// TIA Portal V21 export
// export: Created 2026-11-21T13:31:41.9826464Z, ExportSetting WithDefaults, DisplayName Totally Integrated Automation Portal, DisplayVersion V21, DisplayName STEP 7 Professional, DisplayVersion V21, DisplayName STEP 7 Safety, DisplayVersion V21, DisplayName Tech WebApplication, DisplayVersion V21, DisplayName WinCC Basic/Comfort/Advanced, DisplayVersion V21, DisplayName WinCC Unified, DisplayVersion V21
DATA_BLOCK "Plant"   // DB41
{ S7_Optimized_Access := 'TRUE' }
VERSION : 0.1
// Motors supervised by PlantDiag.
// stored: AutoNumber true, DBAccessibleFromOPCUA true, DBAccessibleFromWebserver true, IsOnlyStoredInLoadMemory false, IsRetainMemResEnabled false, IsWriteProtectedInAS false, MemoryReserve 100
   VAR
      pump : "Motor";
      fans : Array[0..1] of "Motor";
      count : Int;
   END_VAR
BEGIN
END_DATA_BLOCK
